Universal Robots URScript: SplitTest.script

def SplitTest():
  # Global parameters:
  global speed_ms    = 0.250
  global speed_rads  = 0.750
  global accel_mss   = 1.200
  global accel_radss = 1.200
  global blend_radius_m = 0.000

  #--------------------------
  # Add any default subprograms here
  # For example, to drive a gripper as a program call:
  # def Gripper_Open():
  #   ...
  # end
  #
  # Example to drive a spray gun:
  def SprayOn(value):
    # use the value as an output:
    DO_SPRAY = 5
    if value == 0:
      set_standard_digital_out(DO_SPRAY, False)
    else:
      set_standard_digital_out(DO_SPRAY, True)
    end
  end

  # Example to synchronize 2
  def Synchronize():
    # Use the following digital output to signal the state of the robot:
    DO_SYNC = 1

    # Use the following digital input to get the state of another robot:
    DI_SYNC = 1

    if (get_standard_digital_out(DO_SYNC) == get_standard_digital_in(DI_SYNC)):
      set_standard_digital_out(DO_SYNC, not (get_standard_digital_out(DI_SYNC)))
      sleep(0.1)
      thread Thread_wait_1():
        while (True):
          sleep(0.01)
        end
      end
      if (get_standard_digital_out(DO_SYNC) != get_standard_digital_in(DI_SYNC)):
        global thread_handler_1=run Thread_wait_1()
        while (get_standard_digital_out(DO_SYNC) != get_standard_digital_in(DI_SYNC)):
          sync()
        end
        kill thread_handler_1
      end
    else:
      if (get_standard_digital_out(DO_SYNC) != get_standard_digital_in(DI_SYNC)):
        set_standard_digital_out(DO_SYNC, not (get_standard_digital_out(DO_SYNC)))
      end
    end
  end

  #
  # Example to move an external axis
  def MoveAxis(value):
    # use the value as an output:
    DO_AXIS_1 = 1
    DI_AXIS_1 = 1
    if value <= 0:
      set_standard_digital_out(DO_AXIS_1, False)

      # Wait for digital input to change state
      #while (get_standard_digital_in(DI_AXIS_1) != False):
      #  sync()
      #end
    else:
      set_standard_digital_out(DO_AXIS_1, True)

      # Wait for digital input to change state
      #while (get_standard_digital_in(DI_AXIS_1) != True):
      #  sync()
      #end
    end
  end
  #--------------------------


  # Main program:
  # Program generated by VerticalBot Studio for UR5e on 25/10/2026 12:00:00
  # Using nominal kinematics.
  # Using Ref. Frame 2: p[0.100000, -0.050000, 0.020000, 0.000000, 0.000000, 0.523599]
  # set_reference(p[0.100000, -0.050000, 0.020000, 0.000000, 0.000000, 0.523599])
  # Using TCP Tool 1: p[0.010000, 0.000000, 0.120000, 0.000000, 0.261799, 0.000000]
  set_tcp(p[0.010000, 0.000000, 0.120000, 0.000000, 0.261799, 0.000000])
  speed_ms    = 0.2000
  movej([-0.523599, -1.745329, 1.570796, -1.396263, -1.570796, 0.349066],1.20000,0.75000,0,0.0000)
  movel(p[-0.441769, 0.044852, 0.400392, -2.784047, -1.253997, -0.442003],accel_mss,speed_ms,0,0.000)
  movel(p[-0.408198, 0.061237, 0.388074, -2.843025, -1.166595, -0.465806],accel_mss,speed_ms,0,0.000)
  movel(p[-0.441769, 0.044852, 0.400392, -2.784047, -1.253997, -0.442003],accel_mss,speed_ms,0,0.000)
  movel(p[-0.408198, 0.061237, 0.388074, -2.843025, -1.166595, -0.465806],accel_mss,speed_ms,0,0.000)
  movel(p[-0.441769, 0.044852, 0.400392, -2.784047, -1.253997, -0.442003],accel_mss,speed_ms,0,0.000)
  movel(p[-0.408198, 0.061237, 0.388074, -2.843025, -1.166595, -0.465806],accel_mss,speed_ms,0,0.000)
  movel(p[-0.441769, 0.044852, 0.400392, -2.784047, -1.253997, -0.442003],accel_mss,speed_ms,0,0.000)
  movel(p[-0.408198, 0.061237, 0.388074, -2.843025, -1.166595, -0.465806],accel_mss,speed_ms,0,0.000)
  movel(p[-0.441769, 0.044852, 0.400392, -2.784047, -1.253997, -0.442003],accel_mss,speed_ms,0,0.000)
  movel(p[-0.408198, 0.061237, 0.388074, -2.843025, -1.166595, -0.465806],accel_mss,speed_ms,0,0.000)
  movel(p[-0.441769, 0.044852, 0.400392, -2.784047, -1.253997, -0.442003],accel_mss,speed_ms,0,0.000)
  movel(p[-0.408198, 0.061237, 0.388074, -2.843025, -1.166595, -0.465806],accel_mss,speed_ms,0,0.000)
  movel(p[-0.441769, 0.044852, 0.400392, -2.784047, -1.253997, -0.442003],accel_mss,speed_ms,0,0.000)
  movel(p[-0.408198, 0.061237, 0.388074, -2.843025, -1.166595, -0.465806],accel_mss,speed_ms,0,0.000)
  movel(p[-0.441769, 0.044852, 0.400392, -2.784047, -1.253997, -0.442003],accel_mss,speed_ms,0,0.000)
  movel(p[-0.408198, 0.061237, 0.388074, -2.843025, -1.166595, -0.465806],accel_mss,speed_ms,0,0.000)
  movel(p[-0.441769, 0.044852, 0.400392, -2.784047, -1.253997, -0.442003],accel_mss,speed_ms,0,0.000)
  movel(p[-0.408198, 0.061237, 0.388074, -2.843025, -1.166595, -0.465806],accel_mss,speed_ms,0,0.000)
  movel(p[-0.441769, 0.044852, 0.400392, -2.784047, -1.253997, -0.442003],accel_mss,speed_ms,0,0.000)
  movel(p[-0.408198, 0.061237, 0.388074, -2.843025, -1.166595, -0.465806],accel_mss,speed_ms,0,0.000)
  movel(p[-0.441769, 0.044852, 0.400392, -2.784047, -1.253997, -0.442003],accel_mss,speed_ms,0,0.000)
  movel(p[-0.408198, 0.061237, 0.388074, -2.843025, -1.166595, -0.465806],accel_mss,speed_ms,0,0.000)
  movel(p[-0.441769, 0.044852, 0.400392, -2.784047, -1.253997, -0.442003],accel_mss,speed_ms,0,0.000)
  movel(p[-0.408198, 0.061237, 0.388074, -2.843025, -1.166595, -0.465806],accel_mss,speed_ms,0,0.000)
  movel(p[-0.441769, 0.044852, 0.400392, -2.784047, -1.253997, -0.442003],accel_mss,speed_ms,0,0.000)
  movel(p[-0.408198, 0.061237, 0.388074, -2.843025, -1.166595, -0.465806],accel_mss,speed_ms,0,0.000)
  movel(p[-0.441769, 0.044852, 0.400392, -2.784047, -1.253997, -0.442003],accel_mss,speed_ms,0,0.000)
  movel(p[-0.408198, 0.061237, 0.388074, -2.843025, -1.166595, -0.465806],accel_mss,speed_ms,0,0.000)
  movel(p[-0.441769, 0.044852, 0.400392, -2.784047, -1.253997, -0.442003],accel_mss,speed_ms,0,0.000)
  movel(p[-0.408198, 0.061237, 0.388074, -2.843025, -1.166595, -0.465806],accel_mss,speed_ms,0,0.000)
  movel(p[-0.441769, 0.044852, 0.400392, -2.784047, -1.253997, -0.442003],accel_mss,speed_ms,0,0.000)
  movel(p[-0.408198, 0.061237, 0.388074, -2.843025, -1.166595, -0.465806],accel_mss,speed_ms,0,0.000)
  movel(p[-0.441769, 0.044852, 0.400392, -2.784047, -1.253997, -0.442003],accel_mss,speed_ms,0,0.000)
  movel(p[-0.408198, 0.061237, 0.388074, -2.843025, -1.166595, -0.465806],accel_mss,speed_ms,0,0.000)
  movel(p[-0.441769, 0.044852, 0.400392, -2.784047, -1.253997, -0.442003],accel_mss,speed_ms,0,0.000)
  movel(p[-0.408198, 0.061237, 0.388074, -2.843025, -1.166595, -0.465806],accel_mss,speed_ms,0,0.000)
  movel(p[-0.441769, 0.044852, 0.400392, -2.784047, -1.253997, -0.442003],accel_mss,speed_ms,0,0.000)
  movel(p[-0.408198, 0.061237, 0.388074, -2.843025, -1.166595, -0.465806],accel_mss,speed_ms,0,0.000)
  movel(p[-0.441769, 0.044852, 0.400392, -2.784047, -1.253997, -0.442003],accel_mss,speed_ms,0,0.000)
  movel(p[-0.408198, 0.061237, 0.388074, -2.843025, -1.166595, -0.465806],accel_mss,speed_ms,0,0.000)
end

SplitTest()
